# EPICS autosave request: soft_iocs/sydor_bsharp/iocBoot/iocsydor_bsharp_chutch/auto_settings.req
file "quadEM_settings.req",            P=$(P), R=$(R)
